Fanuc KAREL source: KT00456.KL

PROGRAM KT00456
%NOLOCKGROUP
VAR
  P1: POSITION
  P2: XYZWPR
  OUT: BOOLEAN
BEGIN
    P2.Y = 2.0
  OUT = P1 >= P2
END KT00456
